PROGRAM MAIN_Line
VAR
    conveyors : ARRAY[1..3] OF FB_Conveyor;
    motors : ARRAY[1..3] OF FB_MotorSim;
    initialized : BOOL;
    i : DINT;
END_VAR

IF NOT initialized THEN
    FOR i := LOWER_BOUND(conveyors, 1) TO UPPER_BOUND(conveyors, 1) DO
        conveyors[i].BindMotor(motor := motors[i]);
    END_FOR;
    initialized := TRUE;
END_IF;
FOR i := LOWER_BOUND(conveyors, 1) TO UPPER_BOUND(conveyors, 1) DO
    IF GVL_Line.start[i] THEN
        conveyors[i].Start(delay := GVL_Line.startDelay[i]);
    END_IF;
    conveyors[i].Update(guardClosed := GVL_Line.guardClosed[i],
                        stopRequested := GVL_Line.stop[i],
                        sensor := GVL_Line.productSensor[i]);
    GVL_Line.running[i] := conveyors[i].Running;
    GVL_Line.actualSpeed[i] := conveyors[i].ActiveSpeed;
    GVL_Line.productCount[i] := conveyors[i].ProductCount;
    GVL_Line.alarm[i] := conveyors[i].Alarm;
END_FOR;

END_PROGRAM

(* stored: Version 1.1.0.1, ProductVersion 3.1 *)
